// TIA Portal V20 export
// export: Created 2026-10-20T18:54:49.9582785Z, ExportSetting None, DisplayName Totally Integrated Automation Portal, DisplayVersion V20 Update 6, DisplayName TIA Portal Openness, DisplayVersion V20 Update 6, DisplayName TIA Portal Version Control Interface, DisplayVersion V20 Update 6, DisplayName SINAMICS Startdrive Advanced, DisplayVersion V20 SP1, DisplayName SINAMICS Startdrive G130, G150, S120, S150, SINAMICS MV, G220, S200, S210, DisplayVersion V20 SP1, DisplayName SINAMICS Startdrive G110M, G120, G120C, G120D, G120P, G115D, DisplayVersion V20 SP1, DisplayName STEP 7 Professional, DisplayVersion V20 Update 6, DisplayName STEP 7 Safety, DisplayVersion V20 Update 2, DisplayName WinCC Basic/Comfort/Advanced, DisplayVersion V20 Update 6, DisplayName WinCC Unified, DisplayVersion V20 Update 6
VAR_GLOBAL   // PLC tag table "IO_Remote_Panel_2"
   "VTD2 UPPER LIMIT" AT %I164.0 : Bool;
   "VTD2 LOWER LIMIT" AT %I164.3 : Bool;
   "VTD2 PUSH TO ENTER VTD ZONE" AT %I165.4 : Bool;
   "VTD2 PUSH TO EXIT VTD ZONE" AT %I165.5 : Bool;
   "CVTD2 CIRCUIT BREAKER FEEDBACK" AT %I168.0 : Bool;
   "VTD2 CIRCUIT BREAKER FEEDBACK" AT %I168.1 : Bool;
   "CABINET 24V PSU CIRCUIT BREAKER FEEDBACK(2)" AT %I168.2 : Bool;
   "CABINET COOLING FAN CIRCUIT BREAKER FEEDBACK(2)" AT %I168.3 : Bool;
   "OVERTRAVEL LOWER LIMIT - CH1(2)" AT %I558.0 : Bool;   // Overtravel Lower Limit - CH1
   "OVERTRAVEL UPPER LIMIT - CH1(2)" AT %I558.1 : Bool;   // Overtravel Upper Limit - CH1
   "E-STOP (CABINET) - CH1(2)" AT %I558.2 : Bool;   // E-Stop (Cabinet)- CH1
   "RESET (CABINET)(2)" AT %I558.3 : Bool;   // Reset (Cabinet) - CH1
   "OVERTRAVEL LOWER LIMIT - CH2(2)" AT %I558.4 : Bool;   // Overtravel Lower Limit - CH2
   "OVERTRAVEL UPPER LIMIT - CH2(2)" AT %I558.5 : Bool;   // Overtravel Upper Limit - CH2
   "E-STOP (CABINET) - CH2(2)" AT %I558.6 : Bool;   // E-Stop (Cabinet) - CH2
   "Power Enable Safety Stopper Conveyors (Level 7,8 - Side1) - CH1(2)" AT %Q302.0 : Bool;
   "Power Enable Safety Stopper Conveyors (Level 7,8 - Side1) - CH2(2)" AT %Q302.1 : Bool;
   "Power Enable Safety Stopper Conveyors (Level 7,8 - Side2) - CH1(2)" AT %Q302.2 : Bool;
   "Power Enable Safety Stopper Conveyors (Level 7,8 - Side2) - CH2(2)" AT %Q302.3 : Bool;
   "VTU HOIST BRAKE SAFETY ENABLE 1(2)" AT %Q302.4 : Bool;
   "VTU HOIST BRAKE SAFETY ENABLE 2(2)" AT %Q302.5 : Bool;
   "Power Enable Safety Stopper Conveyors (Level 1,2,3 - Side1) - CH1(2)" AT %Q598.0 : Bool;
   "Power Enable Safety Stopper Conveyors (Level 1,2,3 - Side1) - CH2(2)" AT %Q598.1 : Bool;
   "Power Enable Safety Stopper Conveyors (Level 1,2,3 - Side2) - CH1(2)" AT %Q598.2 : Bool;
   "Power Enable Safety Stopper Conveyors (Level 1,2,3 - Side2) - CH2(2)" AT %Q598.3 : Bool;
   "Power Enable Safety Stopper Conveyors (Level 4,5,6 - Side1) - CH1(2)" AT %Q598.4 : Bool;
   "Power Enable Safety Stopper Conveyors (Level 4,5,6 - Side1) - CH2(2)" AT %Q598.5 : Bool;
   "Power Enable Safety Stopper Conveyors (Level 4,5,6 - Side2) - CH1(2)" AT %Q598.6 : Bool;
   "Power Enable Safety Stopper Conveyors (Level 4,5,6 - Side2) - CH2(2)" AT %Q598.7 : Bool;
   "STO VTD - CH1(2)" AT %Q586.0 : Bool;
   "STO VTD - CH2(2)" AT %Q586.1 : Bool;
   "STO CONVEYOR VTD - CH1(2)" AT %Q586.2 : Bool;
   "STO CONVEYOR VTD - CH2(2)" AT %Q586.3 : Bool;
   "STO CNV VFD (Level 1,2,3 - Side1) - CH1(2)" AT %Q586.4 : Bool;
   "STO CNV VFD (Level 1,2,3 - Side1) - CH2(2)" AT %Q586.5 : Bool;
   "STO CNV VFD (Level 1,2,3 - Side2) - CH1(2)" AT %Q586.6 : Bool;
   "STO CNV VFD (Level 1,2,3 - Side2) - CH2(2)" AT %Q586.7 : Bool;
   "STO CNV VFD (Level 4,5,6 - Side1) - CH1(2)" AT %Q592.0 : Bool;
   "STO CNV VFD (Level 4,5,6 - Side1) - CH2(2)" AT %Q592.1 : Bool;
   "STO CNV VFD (Level 4,5,6 - Side2) - CH1(2)" AT %Q592.2 : Bool;
   "STO CNV VFD (Level 4,5,6 - Side2) - CH2(2)" AT %Q592.3 : Bool;
   "STO CNV VFD (Level 7,8 - Side1) - CH1(2)" AT %Q592.4 : Bool;
   "STO CNV VFD (Level 7,8 - Side1) - CH2(2)" AT %Q592.5 : Bool;
   "STO CNV VFD (Level 7,8 - Side2) - CH1(2)" AT %Q592.6 : Bool;
   "STO CNV VFD (Level 7,8 - Side2) - CH2(2)" AT %Q592.7 : Bool;
   "VTD2 SFTY STOPPER CNVS 7,8 - (SIDE 1)" AT %I572.4 : Bool;
   "VTD2 SFTY STOPPER CNVS 1,2,3 - (SIDE 2)" AT %I572.1 : Bool;
   "VTD2 SFTY STOPPER CNVS 1,2,3 - (SIDE 1)" AT %I572.0 : Bool;   // SAFETY STOPPER CONVEYORS (1,2,3 - SIDE 1) EDMFEEDBACK
   "VTU HOIST BRAKE SAFETY ENABLE EDM FEEDBACK(2)" AT %I572.6 : Bool;
   "VTD2 SFTY STOPPER CNVS 4,5,6 - (SIDE 1)" AT %I572.2 : Bool;
   "VTD2 SFTY STOPPER CNVS 7,8 - (SIDE 2)" AT %I572.5 : Bool;
   "EMERGENCY STOP RESET STATUS - ON(2)" AT %Q206.7 : Bool;   // 920SL1
   "VTD2 SFTY STOPPER CNVS 4,5,6 - (SIDE 2)" AT %I572.3 : Bool;
   "C2202 CIRCUIT BREAKER FEEDBACK" AT %I166.1 : Bool;
   "C2106 CIRCUIT BREAKER FEEDBACK" AT %I167.5 : Bool;
   "C2102 CIRCUIT BREAKER FEEDBACK" AT %I167.1 : Bool;
   "C2203 CIRCUIT BREAKER FEEDBACK" AT %I166.2 : Bool;
   "C2107 CIRCUIT BREAKER FEEDBACK" AT %I167.6 : Bool;
   "C2208 CIRCUIT BREAKER FEEDBACK" AT %I166.7 : Bool;
   "C2205 CIRCUIT BREAKER FEEDBACK" AT %I166.4 : Bool;
   "C2206 CIRCUIT BREAKER FEEDBACK" AT %I166.5 : Bool;
   "C2108 CIRCUIT BREAKER FEEDBACK" AT %I167.7 : Bool;
   "C2105 CIRCUIT BREAKER FEEDBACK" AT %I167.4 : Bool;
   "C2204 CIRCUIT BREAKER FEEDBACK" AT %I166.3 : Bool;
   "C2101 CIRCUIT BREAKER FEEDBACK" AT %I167.0 : Bool;
   "C2201 CIRCUIT BREAKER FEEDBACK" AT %I166.0 : Bool;
   "C2103 CIRCUIT BREAKER FEEDBACK" AT %I167.2 : Bool;
   "C2104 CIRCUIT BREAKER FEEDBACK" AT %I167.3 : Bool;
   "C2207 CIRCUIT BREAKER FEEDBACK" AT %I166.6 : Bool;
   "SCA 2002 STACK LIGHTS GREEN" AT %Q206.6 : Bool;
   "C2202_SFTY STOPPER ROTATE" AT %Q198.4 : Bool;
   "C2104_SFTY STOPPER ROTATE" AT %Q203.4 : Bool;
   "C2103_SFTY STOPPER ROTATE" AT %Q203.0 : Bool;
   "C2102_SFTY STOPPER ROTATE" AT %Q202.4 : Bool;
   "C2203_SFTY STOPPER ROTATE" AT %Q199.0 : Bool;
   "C2204_SFTY STOPPER ROTATE" AT %Q199.4 : Bool;
   "C2101_SFTY STOPPER ROTATE" AT %Q202.0 : Bool;
   "C2105_SFTY STOPPER ROTATE" AT %Q204.0 : Bool;
   "C2205_SFTY STOPPER ROTATE" AT %Q200.0 : Bool;
   "C2208_SFTY STOPPER ROTATE" AT %Q201.4 : Bool;
   "C2206_SFTY STOPPER ROTATE" AT %Q200.4 : Bool;
   "C2207_SFTY STOPPER ROTATE" AT %Q201.0 : Bool;
   "C2108_SFTY STOPPER ROTATE" AT %Q205.4 : Bool;
   "C2201_SFTY STOPPER ROTATE" AT %Q198.0 : Bool;
   "C2107_SFTY STOPPER ROTATE" AT %Q205.0 : Bool;
   "C2106_SFTY STOPPER ROTATE" AT %Q204.4 : Bool;
   "Chain Slack 3 - CH1(2)" AT %I565.1 : Bool;   // Chain Slack 3 - CH1
   "Chain Slack 4 - CH2(2)" AT %I565.4 : Bool;   // Chain Slack 4 - CH2
   "Chain Slack 1 - CH1(2)" AT %I565.2 : Bool;   // Chain Slack 1 - CH1
   "Chain Slack 2 - CH2(2)" AT %I565.7 : Bool;   // Chain Slack 2 - CH2
   "Chain Slack 3 - CH2(2)" AT %I565.5 : Bool;   // Chain Slack 3 - CH2
   "SCA 2002 STACK LIGHTS AMBER" AT %Q206.5 : Bool;
   "SCA 2002 STACK LIGHTS RED" AT %Q206.4 : Bool;
   "Chain Slack 4 - CH1(2)" AT %I565.0 : Bool;   // Chain Slack 4 - CH1
   "Chain Slack 1 - CH2(2)" AT %I565.6 : Bool;   // Chain Slack 1 - CH2
   "Chain Slack 2 - CH1(2)" AT %I565.3 : Bool;   // Chain Slack 2 - CH1
   "VTD2 DOCKING PINS 1 EXTEND" AT %Q206.2 : Bool;
   "VTD2 DOCKING PINS 1 RETRACT" AT %Q206.3 : Bool;
   "VTD2 DOCKING PINS 2 EXTEND" AT %Q206.0 : Bool;
   "VTD2 DOCKING PINS 2 RETRACT" AT %Q206.1 : Bool;
   "LIGHT GUARDS C2101 - CH1" AT %I579.1 : Bool;
   "LIGHT GUARDS C2101 - CH2" AT %I579.5 : Bool;
   "LIGHT GUARDS C2201 - CH1" AT %I579.0 : Bool;
   "LIGHT GUARDS C2201 - CH2" AT %I579.4 : Bool;
   "GATE_SENSOR_1_CH1(2)" AT %I579.2 : Bool;
   "GATE_SENSOR_1_CH2(2)" AT %I579.6 : Bool;
   "GATE_SENSOR_2_CH1(2)" AT %I579.3 : Bool;
   "GATE_SENSOR_2_CH2(2)" AT %I579.7 : Bool;
END_VAR
